(* LS Electric XG5000 project: MPST *)
(* PLC LSPLC *)
(* module base 0 slot 0: 입출력 모듈:XEM-DN/DP32HP (DC 24V 입력, 트랜지스터 출력 32점 (싱크출력/소스출력)) *)
(* module base 0 slot 1: 내장위치결정:XBF-PO06E (오픈컬렉터형, 6축) *)

PROGRAM NewProgram (* task: 스캔 프로그램 *)
VAR
    Count : INT; (* Source preservation check *)
END_VAR
Count := Count + 1;
END_PROGRAM

PROGRAM AddedST (* task: 스캔 프로그램 *)
VAR
    Count : INT; (* Source preservation check *)
END_VAR
Count := Count + 1;
END_PROGRAM

PROGRAM AddedIL (* task: 스캔 프로그램 *)
VAR
    Count : INT; (* Source preservation check *)
END_VAR
LD Count
ADD 1
ST Count
END_PROGRAM